(* PLC project VoltPilot-Vorlage PV, VoltPilot VoltPilot EMS 1.0 *)
(* stored: creationDateTime 2026-11-20T00:00:00 *)

(* VoltPilot-Bibliothek · Datentypen des Bausteins Erzeuger-Bild Das Anlagenprogramm füllt diese Strukturen in den Einheiten der Felder des Vertrags docs/contracts/v2/erzeuger-registerbild.md (W, kW, 0,1 %, 0,001, 0,1 kWh, s) und rechnet keine Register: das tut FB_VP_ErzeugerBild. Ein Wert ohne deckendes Gültigkeitsbit hat ein eigenes Feld ...Bekannt: FALSE heißt "kein Wert", der Baustein schreibt dann das Typ-Maximum (Vertrag §1: ungültig ist nie 0). Ein gedeckter Wert braucht keines: ist sein Gültigkeitsbit FALSE, schreibt der Baustein das Typ-Maximum selbst. Ausnahme ist uiPZehntelProzent (Vertrag §3, Wort 24): ohne gültige Vorgabe steht dort der wirksame Ersatzwert. Das Eingangsregister-Abbild: Bild 0..137, Namen ab 140 (höchstens 140 + 32 + 16 * 10 = 332 Wörter). *)
TYPE T_VP_ErzeugerBild : ARRAY[0..331] OF WORD;
END_TYPE

(* Abschnitt A: Anlage und Netzpunkt (Register 12..21). *)
TYPE ST_VP_ErzeugerAnlage : STRUCT
  xNetzpunktGueltig : BOOL;
  xNetzpunktBerechnet : BOOL;
  xNetzpunktTot : BOOL;
  xErzeugungGueltig : BOOL;
  xGasspeicherGueltig : BOOL;
  xGueltigBekannt : BOOL := TRUE;
  uiAlterS : UINT;
  xAlterBekannt : BOOL := TRUE;
  diPNetzpunktW : DINT;
  diPErzeugungW : DINT;
  uiZustand : UINT;
  xZustandBekannt : BOOL := TRUE;
  xNotAus : BOOL;
  xNaSchutz : BOOL;
  xSammelstoerung : BOOL;
  xHandOrt : BOOL;
  xWartung : BOOL;
  xBitsBekannt : BOOL := TRUE;
  uiSpeicherZehntelProzent : UINT;
  uiInstalliertKw : UINT;
  xInstalliertBekannt : BOOL := TRUE;
END_STRUCT;
END_TYPE

(* Abschnitt N: Netzbetreiber (Register 22..27). *)
TYPE ST_VP_ErzeugerNetzbetreiber : STRUCT
  uiKanal : UINT;
  xKanalBekannt : BOOL := TRUE;
  xVorgabeGueltig : BOOL;
  xVerbindungSteht : BOOL;
  xWirkleistungBegrenzt : BOOL;
  xNotAus : BOOL;
  xCosPhiVorgabe : BOOL;
  xKennlinie : BOOL;
  xBitsBekannt : BOOL := TRUE;
  uiPZehntelProzent : UINT;
  xPBekannt : BOOL := TRUE;
  iCosPhiTausendstel : INT;
  uiSeitS : UINT;
  xSeitBekannt : BOOL := TRUE;
  uiZaehler : UINT;
END_STRUCT;
END_TYPE

(* Abschnitt D: Direktvermarkter (Register 28..33). *)
TYPE ST_VP_ErzeugerDirektvermarkter : STRUCT
  uiKanal : UINT;
  xKanalBekannt : BOOL := TRUE;
  xAbschnittGueltig : BOOL;
  xAktivierung : BOOL;
  xStopp : BOOL;
  xBereitGemeldet : BOOL;
  xAktivGemeldet : BOOL;
  xBitsBekannt : BOOL := TRUE;
  udiSollW : UDINT;
  uiSeitS : UINT;
  uiZaehler : UINT;
END_STRUCT;
END_TYPE

(* Abschnitt S: Wirkung (Register 34..37). *)
TYPE ST_VP_ErzeugerWirkung : STRUCT
  xGueltig : BOOL;
  xAnlageFolgt : BOOL;
  xBitsBekannt : BOOL := TRUE;
  uiQuelle : UINT;
  udiGrenzeW : UDINT;
END_STRUCT;
END_TYPE

(* Abschnitt T: eine Einheit (Wechselrichter oder BHKW-Motor), 10 Wörter ab 38 + (n - 1) * 10. *)
TYPE ST_VP_ErzeugerEinheit : STRUCT
  xWerteGueltig : BOOL;
  xSollwertGueltig : BOOL;
  xDvBereit : BOOL;
  xDvAktiv : BOOL;
  xGrundStoerung : BOOL;
  xGrundNetzbetreiber : BOOL;
  xGrundHandOrt : BOOL;
  xGrundWartung : BOOL;
  xGrundGasspeicherLeer : BOOL;
  xGrundSonstiger : BOOL;
  xBitsBekannt : BOOL := TRUE;
  uiZustand : UINT;
  uiArt : UINT;
  xArtBekannt : BOOL := TRUE;
  uiNennKw : UINT;
  xNennBekannt : BOOL := TRUE;
  diPIstW : DINT;
  udiPSollW : UDINT;
  udiEZehntelKwh : UDINT;
  sTyp : STRING(32);
END_STRUCT;
END_TYPE

(* VoltPilot-Bibliothek · Datentypen des Koppelbilds (docs/contracts/v2/koppelbild.md) Das Anlagenprogramm sieht keine Register: es trägt je Stellplatz ein Angebot ein, liest den Wunsch am Ausgang des Bausteins und meldet zurück, was es wirklich anwendet. Codes (Vertrag §7): Art 0 keiner, 1 limit_w (W), 2 limit_pct (0,1 %), 3 setpoint_w (W, Speicher + lädt), 4 on_off (0/1), 5 mode (1..8), 6 setpoint_c (0,1 °C) Ziel 1 erzeugung_gesamt, 2 erzeugungseinheit, 3 speicher, 4 verbraucher, 5 netzbezug, 6 einspeisung, 7 probe Grund 0 keiner, 1 markt, 2 netz, 3 regel, 4 hand, 5 test, 6 vertrag (Nebenversion 1.1; Auskunft, keine Weiche: der Baustein reicht ihn unverändert durch) Abschnitt W: liegt auf den Halteregistern 0..63 des Modbus-TCP-Servers; nur die Edge schreibt. *)
TYPE T_VP_KoppelWunsch : ARRAY[0..63] OF WORD;
END_TYPE

(* Abschnitt Q: liegt auf den Eingangsregistern 1000..1115; nur der Baustein schreibt. *)
TYPE T_VP_KoppelQuittung : ARRAY[0..115] OF WORD;
END_TYPE

(* Was ein Stellplatz anbietet. uiArt 0 = Platz leer. Band in den Einheiten der Art. *)
TYPE ST_VP_Angebot : STRUCT
  uiArt : UINT;
  uiZiel : UINT;
  uiNr : UINT;
  diMin : DINT;
  diMax : DINT;
  xBereit : BOOL;
  xGrundStoerung : BOOL;
  xGrundHandOrt : BOOL;
  xGrundWartung : BOOL;
  xGrundVorrang : BOOL;
  xGrundSonstiger : BOOL;
END_STRUCT;
END_TYPE

(* Was das Anlagenprogramm für das Ziel eines Stellplatzes gerade anwendet, gleich woher es kommt. *)
TYPE ST_VP_Rueckmeldung : STRUCT
  diWirksam : DINT;
  xWirksamBekannt : BOOL;
  xUeberstimmt : BOOL;
END_STRUCT;
END_TYPE

(* Der zugelassene Wunsch eines Stellplatzes. Ohne xGilt fährt das Anlagenprogramm mit eigenen Werten. *)
TYPE ST_VP_Wunsch : STRUCT
  xGilt : BOOL;
  diWert : DINT;
  uiGrund : UINT;
  uiUrteil : UINT;
END_STRUCT;
END_TYPE

(* VoltPilot-Bibliothek · Datentypen des Bausteins WAGO-Bild (Energiekarten) Das Anlagenprogramm kopiert je 3-Phasen-Leistungsmessklemme 750-494/-495 („Energiekarte“) die Werte, die es aus der Karte gelesen hat, in eine ST_VP_WagoKarte - unverändert, in der Skalierung der Karte (docs/contracts/v2/wago-registerbild.md §4). Umgerechnet wird nichts: Einheit, Faktor und Vorzeichen kommen aus dem Katalog und dem Hardwareblatt der Anlage. Jeder Teil hat sein Feld ...Gelesen: FALSE heißt "dieser Teil ist unbekannt", der Baustein löscht dann das Gültigkeitsbit und schreibt das Typ-Maximum - nie 0, nie einen alten Wert. Das Abbild: Kopf 12 Wörter und höchstens 16 Karten zu je 42 Wörtern (12 + 16 * 42 = 684). *)
TYPE T_VP_WagoBild : ARRAY[0..683] OF WORD;
END_TYPE

(* Eine Energiekarte (Vertrag §4). *)
TYPE ST_VP_WagoKarte : STRUCT
  uiSteckplatz : UINT;
  uiKartentyp : UINT;
  uiVariante : UINT;
  xKarteGelesen : BOOL;
  xKr32Gelesen : BOOL;
  wKr32 : WORD;
  xKr35Gelesen : BOOL;
  wKr35 : WORD;
  xStatusGelesen : BOOL;
  awStatus : ARRAY[0..11] OF WORD;
  adwMesswert : ARRAY[1..12] OF DWORD;
END_STRUCT;
END_TYPE

VAR_GLOBAL  (* GVL_VoltPilot *)
  aErzeugerBild : T_VP_ErzeugerBild;
  aKoppelQuittung : T_VP_KoppelQuittung;
  aKoppelWunsch : T_VP_KoppelWunsch;
  aWagoBild : T_VP_WagoBild;
  xProbeLampe : BOOL;
END_VAR

(* VoltPilot-Bibliothek · Baustein Erzeuger-Bild Füllt das "VoltPilot-Registerbild Erzeuger v1" (schlanke Fassung 1.0, docs/contracts/v2/erzeuger-registerbild.md) aus den getippten Werten des Anlagenprogramms. Das Abbild aBild liegt auf den Eingangsregistern des Modbus-TCP-Servers ab Adresse 0 (Funktionscode 4); die Box liest es alle 5 s, auf einem PFC200 mit VoltPilot über 127.0.0.1. Aufruf: einmal je Zyklus in der Task, die das Abbild auch dem Modbus-Server übergibt. fbBild(uiProgrammstand := 2611, uiAnlagenart := 1, uiTeAnzahl := 3, stAnlage := stAnlage, stNetzbetreiber := stNb, stDirektvermarkter := stDv, stWirkung := stWirkung, astEinheit := astEinheit, xMitNamen := TRUE, sNetzbetreiber := 'Netzbetreiber', sDirektvermarkter := '', aBild := GVL_VoltPilot.aErzeugerBild); Was der Baustein selbst hält: - Kopf: Signatur, Prüfwert, Fassung 1.0 - feste Werte, der Prüfwert über VP_SetzeU32; - Herzschlag: +1 je Sekunde seit Programmstart, 65535 -> 0 (Vertrag §8); bleibt der Aufruf aus, steht er, und die Box hält alle Werte nach drei gleichen Lesungen für veraltet; - Typ-Maximum für jeden gedeckten Wert, dessen Gültigkeitsbit fehlt; - Wörter von Einheiten über uiTeAnzahl hinaus und ohne Namen den Namenbereich auf 0. Grenzen: höchstens 10 Einheiten; uiTeAnzahl 0 oder über 10 schreibt der Baustein, wie er sie bekommt - die Box liest das Bild dann nicht (te_anzahl_ungueltig), sieht aber Kopf und Herzschlag (so meldet sich das Grundprogramm ohne Anlage). *)
FUNCTION_BLOCK FB_VP_ErzeugerBild
  VAR_INPUT
    udiSteuerungId : UDINT := 16#FFFFFFFF;
    uiProgrammstand : UINT := 16#FFFF;
    uiAnlagenart : UINT := 16#FFFF;
    uiTeAnzahl : UINT;
    stAnlage : ST_VP_ErzeugerAnlage;
    stNetzbetreiber : ST_VP_ErzeugerNetzbetreiber;
    stDirektvermarkter : ST_VP_ErzeugerDirektvermarkter;
    stWirkung : ST_VP_ErzeugerWirkung;
    astEinheit : ARRAY[1..10] OF ST_VP_ErzeugerEinheit;
    xMitNamen : BOOL;
    sNetzbetreiber : STRING(32);
    sDirektvermarkter : STRING(32);
  END_VAR
  VAR_IN_OUT
    aBild : T_VP_ErzeugerBild;
  END_VAR
  VAR
    uiHerzschlag : UINT;
    xGestartet : BOOL;
    tLetzte : TIME;
    tJetzt : TIME;
    udiSekunden : UDINT;
    n : UINT;
    uiBasis : UINT;
    i : UINT;
    wBits : WORD;
  END_VAR

(* --- Herzschlag: +1 je Sekunde, beim Programmstart 0, 65535 -> 0 ---------------------------- *)
tJetzt := TIME();
IF NOT xGestartet THEN
    tLetzte := tJetzt;
    xGestartet := TRUE;
END_IF
udiSekunden := TIME_TO_UDINT(tJetzt - tLetzte) / 1000;
IF udiSekunden > 0 THEN
    uiHerzschlag := uiHerzschlag + UDINT_TO_UINT(udiSekunden AND 16#FFFF);
    tLetzte := tLetzte + UDINT_TO_TIME(udiSekunden * 1000);
END_IF

(* --- Kopf (0..11) ------------------------------------------------------------------------- *)
aBild[0] := 16#5650;   (* "VP" *)
aBild[1] := 16#455A;   (* "EZ" *)
VP_SetzeU32(aBild := aBild, uiAdresse := 2, udiWert := 16#01020304, xBekannt := TRUE);
aBild[4] := 16#0100;   (* Fassung 1.0 *)
aBild[5] := UINT_TO_WORD(uiTeAnzahl);
aBild[6] := UINT_TO_WORD(uiHerzschlag);
aBild[7] := UINT_TO_WORD(uiProgrammstand);
VP_SetzeU32(aBild := aBild, uiAdresse := 8, udiWert := udiSteuerungId, xBekannt := TRUE);
aBild[10] := UINT_TO_WORD(uiAnlagenart);
IF xMitNamen THEN
    aBild[11] := 140;
ELSE
    aBild[11] := 0;
END_IF

(* --- A: Anlage und Netzpunkt (12..21) ------------------------------------------------------ *)
wBits := VP_Bit(stAnlage.xNetzpunktGueltig, 0) OR VP_Bit(stAnlage.xNetzpunktBerechnet, 1)
    OR VP_Bit(stAnlage.xNetzpunktTot, 2) OR VP_Bit(stAnlage.xErzeugungGueltig, 3)
    OR VP_Bit(stAnlage.xGasspeicherGueltig, 4);
VP_SetzeU16(aBild := aBild, uiAdresse := 12, uiWert := WORD_TO_UINT(wBits), xBekannt := stAnlage.xGueltigBekannt);
VP_SetzeU16(aBild := aBild, uiAdresse := 13, uiWert := stAnlage.uiAlterS, xBekannt := stAnlage.xAlterBekannt);
VP_SetzeS32(aBild := aBild, uiAdresse := 14, diWert := stAnlage.diPNetzpunktW,
    xBekannt := stAnlage.xGueltigBekannt AND stAnlage.xNetzpunktGueltig);
VP_SetzeS32(aBild := aBild, uiAdresse := 16, diWert := stAnlage.diPErzeugungW,
    xBekannt := stAnlage.xGueltigBekannt AND stAnlage.xErzeugungGueltig);
VP_SetzeU16(aBild := aBild, uiAdresse := 18, uiWert := stAnlage.uiZustand, xBekannt := stAnlage.xZustandBekannt);
wBits := VP_Bit(stAnlage.xNotAus, 0) OR VP_Bit(stAnlage.xNaSchutz, 1) OR VP_Bit(stAnlage.xSammelstoerung, 2)
    OR VP_Bit(stAnlage.xHandOrt, 3) OR VP_Bit(stAnlage.xWartung, 4);
VP_SetzeU16(aBild := aBild, uiAdresse := 19, uiWert := WORD_TO_UINT(wBits), xBekannt := stAnlage.xBitsBekannt);
VP_SetzeU16(aBild := aBild, uiAdresse := 20, uiWert := stAnlage.uiSpeicherZehntelProzent,
    xBekannt := stAnlage.xGueltigBekannt AND stAnlage.xGasspeicherGueltig);
VP_SetzeU16(aBild := aBild, uiAdresse := 21, uiWert := stAnlage.uiInstalliertKw, xBekannt := stAnlage.xInstalliertBekannt);

(* --- N: Netzbetreiber (22..27) ------------------------------------------------------------- *)
VP_SetzeU16(aBild := aBild, uiAdresse := 22, uiWert := stNetzbetreiber.uiKanal, xBekannt := stNetzbetreiber.xKanalBekannt);
wBits := VP_Bit(stNetzbetreiber.xVorgabeGueltig, 0) OR VP_Bit(stNetzbetreiber.xVerbindungSteht, 1)
    OR VP_Bit(stNetzbetreiber.xWirkleistungBegrenzt, 2) OR VP_Bit(stNetzbetreiber.xNotAus, 3)
    OR VP_Bit(stNetzbetreiber.xCosPhiVorgabe, 4) OR VP_Bit(stNetzbetreiber.xKennlinie, 5);
VP_SetzeU16(aBild := aBild, uiAdresse := 23, uiWert := WORD_TO_UINT(wBits), xBekannt := stNetzbetreiber.xBitsBekannt);
(* Wort 24 ohne gültige Vorgabe: der wirksame Ersatzwert, nicht das Typ-Maximum (Vertrag §3) *)
VP_SetzeU16(aBild := aBild, uiAdresse := 24, uiWert := stNetzbetreiber.uiPZehntelProzent, xBekannt := stNetzbetreiber.xPBekannt);
VP_SetzeS16(aBild := aBild, uiAdresse := 25, iWert := stNetzbetreiber.iCosPhiTausendstel,
    xBekannt := stNetzbetreiber.xBitsBekannt AND stNetzbetreiber.xVorgabeGueltig);
VP_SetzeU16(aBild := aBild, uiAdresse := 26, uiWert := stNetzbetreiber.uiSeitS, xBekannt := stNetzbetreiber.xSeitBekannt);
aBild[27] := UINT_TO_WORD(stNetzbetreiber.uiZaehler);

(* --- D: Direktvermarkter (28..33) ---------------------------------------------------------- *)
VP_SetzeU16(aBild := aBild, uiAdresse := 28, uiWert := stDirektvermarkter.uiKanal, xBekannt := stDirektvermarkter.xKanalBekannt);
wBits := VP_Bit(stDirektvermarkter.xAbschnittGueltig, 0) OR VP_Bit(stDirektvermarkter.xAktivierung, 1)
    OR VP_Bit(stDirektvermarkter.xStopp, 2) OR VP_Bit(stDirektvermarkter.xBereitGemeldet, 3)
    OR VP_Bit(stDirektvermarkter.xAktivGemeldet, 4);
VP_SetzeU16(aBild := aBild, uiAdresse := 29, uiWert := WORD_TO_UINT(wBits), xBekannt := stDirektvermarkter.xBitsBekannt);
VP_SetzeU32(aBild := aBild, uiAdresse := 30, udiWert := stDirektvermarkter.udiSollW,
    xBekannt := stDirektvermarkter.xBitsBekannt AND stDirektvermarkter.xAbschnittGueltig);
VP_SetzeU16(aBild := aBild, uiAdresse := 32, uiWert := stDirektvermarkter.uiSeitS,
    xBekannt := stDirektvermarkter.xBitsBekannt AND stDirektvermarkter.xAbschnittGueltig);
(* d_zaehler hat keinen Ungültig-Wert; ohne gültigen Abschnitt liest ihn die Box nicht *)
aBild[33] := UINT_TO_WORD(stDirektvermarkter.uiZaehler);

(* --- S: Wirkung (34..37) ------------------------------------------------------------------- *)
VP_SetzeU16(aBild := aBild, uiAdresse := 34, uiWert := stWirkung.uiQuelle,
    xBekannt := stWirkung.xBitsBekannt AND stWirkung.xGueltig);
wBits := VP_Bit(stWirkung.xGueltig, 0) OR VP_Bit(stWirkung.xAnlageFolgt, 1);
VP_SetzeU16(aBild := aBild, uiAdresse := 35, uiWert := WORD_TO_UINT(wBits), xBekannt := stWirkung.xBitsBekannt);
VP_SetzeU32(aBild := aBild, uiAdresse := 36, udiWert := stWirkung.udiGrenzeW,
    xBekannt := stWirkung.xBitsBekannt AND stWirkung.xGueltig);

(* --- T: je Einheit 10 Wörter ab 38 + (n - 1) * 10 ------------------------------------------ *)
FOR n := 1 TO 10 DO
    uiBasis := 38 + (n - 1) * 10;
    IF n <= uiTeAnzahl THEN
        VP_SetzeU16(aBild := aBild, uiAdresse := uiBasis, uiWert := astEinheit[n].uiZustand,
            xBekannt := astEinheit[n].xBitsBekannt AND astEinheit[n].xWerteGueltig);
        wBits := VP_Bit(astEinheit[n].xWerteGueltig, 0) OR VP_Bit(astEinheit[n].xSollwertGueltig, 1)
            OR VP_Bit(astEinheit[n].xDvBereit, 2) OR VP_Bit(astEinheit[n].xDvAktiv, 3)
            OR VP_Bit(astEinheit[n].xGrundStoerung, 4) OR VP_Bit(astEinheit[n].xGrundNetzbetreiber, 5)
            OR VP_Bit(astEinheit[n].xGrundHandOrt, 6) OR VP_Bit(astEinheit[n].xGrundWartung, 7)
            OR VP_Bit(astEinheit[n].xGrundGasspeicherLeer, 8) OR VP_Bit(astEinheit[n].xGrundSonstiger, 9);
        VP_SetzeU16(aBild := aBild, uiAdresse := uiBasis + 1, uiWert := WORD_TO_UINT(wBits),
            xBekannt := astEinheit[n].xBitsBekannt);
        VP_SetzeU16(aBild := aBild, uiAdresse := uiBasis + 2, uiWert := astEinheit[n].uiArt,
            xBekannt := astEinheit[n].xArtBekannt);
        VP_SetzeU16(aBild := aBild, uiAdresse := uiBasis + 3, uiWert := astEinheit[n].uiNennKw,
            xBekannt := astEinheit[n].xNennBekannt);
        VP_SetzeS32(aBild := aBild, uiAdresse := uiBasis + 4, diWert := astEinheit[n].diPIstW,
            xBekannt := astEinheit[n].xBitsBekannt AND astEinheit[n].xWerteGueltig);
        VP_SetzeU32(aBild := aBild, uiAdresse := uiBasis + 6, udiWert := astEinheit[n].udiPSollW,
            xBekannt := astEinheit[n].xBitsBekannt AND astEinheit[n].xSollwertGueltig);
        VP_SetzeU32(aBild := aBild, uiAdresse := uiBasis + 8, udiWert := astEinheit[n].udiEZehntelKwh,
            xBekannt := astEinheit[n].xBitsBekannt AND astEinheit[n].xWerteGueltig);
    ELSE
        (* frei: nichts Altes aus einer früheren Zahl der Einheiten bleibt stehen *)
        FOR i := uiBasis TO uiBasis + 9 DO
            aBild[i] := 0;
        END_FOR
    END_IF
END_FOR
FOR i := 138 TO 139 DO
    aBild[i] := 0;
END_FOR

(* --- Namen ab 140: Netzbetreiber +0, Direktvermarkter +16, Typ der Einheit n +32 + (n - 1) * 16 *)
IF xMitNamen THEN
    VP_SetzeText(aBild := aBild, uiAdresse := 140, sText := sNetzbetreiber);
    VP_SetzeText(aBild := aBild, uiAdresse := 156, sText := sDirektvermarkter);
    FOR n := 1 TO 10 DO
        IF n <= uiTeAnzahl THEN
            VP_SetzeText(aBild := aBild, uiAdresse := 172 + (n - 1) * 16, sText := astEinheit[n].sTyp);
        ELSE
            VP_SetzeText(aBild := aBild, uiAdresse := 172 + (n - 1) * 16, sText := '');
        END_IF
    END_FOR
ELSE
    FOR i := 140 TO 331 DO
        aBild[i] := 0;
    END_FOR
END_IF
END_FUNCTION_BLOCK

(* VoltPilot-Bibliothek · Baustein Koppelbild Die SPS-Seite des "VoltPilot-Koppelbild v1" (docs/contracts/v2/koppelbild.md): die Edge schreibt Wünsche in die Halteregister 0..63, der Baustein prüft sie, begrenzt jeden auf das Angebot und reicht ihn dem Anlagenprogramm; die Quittung steht in den Eingangsregistern 1000..1115. Die SPS entscheidet immer selbst: ein Wunsch ist nie ein Befehl. Aufruf: einmal je Zyklus in der Task, die die Abbilder auch dem Modbus-Server übergibt. fbKoppel(udiSteuerungId := 1042, xFernsteuerungFrei := xSchluesselFern, xHandOrt := xHand, aAngebot := aAngebot, aRueckmeldung := aRueck, aWunschRegister := GVL_VoltPilot.aKoppelWunsch, aQuittungRegister := GVL_VoltPilot.aKoppelQuittung); IF fbKoppel.aWunsch[1].xGilt THEN diGrenze := MIN(diGrenze, fbKoppel.aWunsch[1].diWert); END_IF Was der Baustein selbst hält: - jeder Wunsch läuft von selbst ab: höchstens frist_s ab Empfang, nie länger als tHoechsteFrist (Vorgabe 60 s); fällt die Edge aus, fährt die Anlage danach mit eigenen Werten; - Lebenszeichen: Herzschlag +1 je Sekunde (wie im Erzeuger-Bild), edge_lebt aus dem letzten gültigen Telegramm; - geprüft wird nur ein Telegramm, dessen Wörter sich geändert haben, in der Reihenfolge von Vertrag §5; ein abgelehntes bewirkt nichts, das vorige gilt bis zu seiner Frist; - Hand/Ort nimmt jedem Stellplatz die Bereitschaft; ohne Fernsteuerung gilt kein Wunsch. Was beim ersten Aufruf in den Halteregistern steht, ist kein Telegramm, nur der Vergleichsstand. *)
FUNCTION_BLOCK FB_VP_Koppelbild
  VAR_INPUT
    udiSteuerungId : UDINT;
    xFernsteuerungFrei : BOOL;
    xHandOrt : BOOL;
    aAngebot : ARRAY[1..8] OF ST_VP_Angebot;
    aRueckmeldung : ARRAY[1..8] OF ST_VP_Rueckmeldung;
    tHoechsteFrist : TIME := T#60S;
    uiBibliothek : UINT := 16#0100;
  END_VAR
  VAR_OUTPUT
    aWunsch : ARRAY[1..8] OF ST_VP_Wunsch;
    xEdgeLebt : BOOL;
    uiKopfUrteil : UINT;
    uiRestS : UINT;
  END_VAR
  VAR_IN_OUT
    aWunschRegister : T_VP_KoppelWunsch;
    aQuittungRegister : T_VP_KoppelQuittung;
  END_VAR
  VAR
    uiHerzschlag : UINT;
    xGestartet : BOOL;
    tLetzte : TIME;
    tJetzt : TIME;
    udiSekunden : UDINT;
    xErster : BOOL := TRUE;
    aLetzte : T_VP_KoppelWunsch;
    aGilt : T_VP_KoppelWunsch;
    xHatTelegramm : BOOL;
    xFristLaeuft : BOOL;
    uiOhneFrist : UINT;
    tAnnahme : TIME;
    udiFristMs : UDINT;
    udiSeitMs : UDINT;
    xLebt : BOOL;
    uiQSitzung : UINT;
    uiQHerzschlag : UINT;
    uiAngenommen : UINT;
    uiAbgelehnt : UINT;
    xGeaendert : BOOL;
    uiGrund : UINT;
    udiFrist : UDINT;
    i : UINT;
    n : UINT;
    uiW : UINT;
    uiQ : UINT;
    uiAnzahl : UINT;
    xLeer : BOOL;
    xBereit : BOOL;
    uiArtW : UINT;
    diW : DINT;
    diWert : DINT;
    uiUrteil : UINT;
  END_VAR

(* --- Herzschlag: +1 je Sekunde seit Programmstart, 65535 -> 0 ------------------------------ *)
tJetzt := TIME();
IF NOT xGestartet THEN
    tLetzte := tJetzt;
    xGestartet := TRUE;
END_IF
udiSekunden := TIME_TO_UDINT(tJetzt - tLetzte) / 1000;
IF udiSekunden > 0 THEN
    uiHerzschlag := uiHerzschlag + UDINT_TO_UINT(udiSekunden AND 16#FFFF);
    tLetzte := tLetzte + UDINT_TO_TIME(udiSekunden * 1000);
END_IF

(* --- Telegramm prüfen, wenn sich ein Wort geändert hat (Vertrag §5) ------------------------- *)
IF xErster THEN
    aLetzte := aWunschRegister;
    xErster := FALSE;
ELSE
    xGeaendert := FALSE;
    FOR i := 0 TO 63 DO
        IF aWunschRegister[i] <> aLetzte[i] THEN
            xGeaendert := TRUE;
        END_IF
    END_FOR
    IF xGeaendert THEN
        aLetzte := aWunschRegister;
        udiFrist := WORD_TO_UDINT(aWunschRegister[10]);
        uiGrund := 0;
        IF aWunschRegister[0] <> 16#5650 OR aWunschRegister[1] <> 16#4B57 THEN
            uiGrund := 2;
        ELSIF SHR(aWunschRegister[4], 8) <> 1 THEN
            uiGrund := 3;
        ELSIF aWunschRegister[2] <> 16#0102 OR aWunschRegister[3] <> 16#0304 THEN
            uiGrund := 4;
        ELSIF VP_KoppelSiegelW(aW := aWunschRegister) <> aWunschRegister[15] THEN
            uiGrund := 5;
        ELSIF VP_KoppelLiesU32(aW := aWunschRegister, uiAdresse := 8) <> udiSteuerungId THEN
            uiGrund := 6;
        ELSIF udiFrist < 5 OR udiFrist > 600 OR aWunschRegister[6] = 0 OR aWunschRegister[6] = 16#FFFF
                OR aWunschRegister[5] <> 8 THEN
            uiGrund := 7;
        END_IF
        IF uiGrund <> 0 THEN
            (* dieses Telegramm bewirkt nichts; das vorige gilt bis zu seiner Frist *)
            uiAbgelehnt := uiAbgelehnt + 1;
            uiKopfUrteil := uiGrund;
        ELSE
            aGilt := aWunschRegister;
            xHatTelegramm := TRUE;
            uiQSitzung := WORD_TO_UINT(aWunschRegister[6]);
            uiQHerzschlag := WORD_TO_UINT(aWunschRegister[7]);
            uiAngenommen := uiAngenommen + 1;
            tAnnahme := tJetzt;
            xLebt := TRUE;
            IF xFernsteuerungFrei THEN
                udiFristMs := MIN(udiFrist * 1000, TIME_TO_UDINT(tHoechsteFrist));
                xFristLaeuft := TRUE;
                uiKopfUrteil := 1;
            ELSE
                xFristLaeuft := FALSE;
                uiOhneFrist := 2;
                uiKopfUrteil := 9;
            END_IF
        END_IF
    END_IF
END_IF

(* --- Fernsteuerung entzogen: alle Wünsche fallen sofort ------------------------------------ *)
IF NOT xFernsteuerungFrei AND xFristLaeuft THEN
    xFristLaeuft := FALSE;
    uiOhneFrist := 2;
    uiKopfUrteil := 9;
END_IF

(* --- Frist: läuft von selbst ab ------------------------------------------------------------ *)
udiSeitMs := TIME_TO_UDINT(tJetzt - tAnnahme);
IF xFristLaeuft AND udiSeitMs >= udiFristMs THEN
    xFristLaeuft := FALSE;
    uiOhneFrist := 1;
    uiKopfUrteil := 8;
END_IF
IF xFristLaeuft THEN
    uiRestS := UDINT_TO_UINT((udiFristMs - udiSeitMs + 999) / 1000);
ELSE
    uiRestS := 0;
END_IF
(* einmal still, bleibt still: auch wenn TIME() nach 49 Tagen überläuft *)
IF xLebt AND udiSeitMs >= 15000 THEN
    xLebt := FALSE;
END_IF
xEdgeLebt := xLebt;

(* --- Kopf der Quittung (1000..1019, hier 0..19) -------------------------------------------- *)
aQuittungRegister[0] := 16#5650;   (* "VP" *)
aQuittungRegister[1] := 16#4B51;   (* "KQ" *)
VP_KoppelSetzeU32(aQ := aQuittungRegister, uiAdresse := 2, udiWert := 16#01020304);
aQuittungRegister[4] := 16#0100;   (* Fassung 1.0 *)
aQuittungRegister[6] := UINT_TO_WORD(uiHerzschlag);
aQuittungRegister[7] := UINT_TO_WORD(uiBibliothek);
VP_KoppelSetzeU32(aQ := aQuittungRegister, uiAdresse := 8, udiWert := udiSteuerungId);
aQuittungRegister[10] := UINT_TO_WORD(uiKopfUrteil);
aQuittungRegister[11] := UINT_TO_WORD(uiQSitzung);
aQuittungRegister[12] := UINT_TO_WORD(uiQHerzschlag);
aQuittungRegister[13] := UINT_TO_WORD(uiRestS);
aQuittungRegister[14] := VP_Bit(xGesetzt := xFernsteuerungFrei, uiBit := 0)
    OR VP_Bit(xGesetzt := xLebt, uiBit := 1) OR VP_Bit(xGesetzt := xHandOrt, uiBit := 2);
aQuittungRegister[15] := UINT_TO_WORD(uiAngenommen);
aQuittungRegister[16] := UINT_TO_WORD(uiAbgelehnt);
aQuittungRegister[17] := 0;
aQuittungRegister[18] := 0;

(* --- je Stellplatz: Angebot, Urteil, zugelassener Wert, wirksam (Vertrag §5) ---------------- *)
uiAnzahl := 0;
FOR n := 1 TO 8 DO
    uiW := 16 + (n - 1) * 6;
    uiQ := 20 + (n - 1) * 12;
    xLeer := aAngebot[n].uiArt = 0;
    xBereit := NOT xLeer AND aAngebot[n].xBereit AND NOT xHandOrt;
    uiUrteil := 0;
    diWert := 0;
    aWunsch[n].xGilt := FALSE;
    aWunsch[n].uiGrund := 0;
    IF NOT xLeer THEN
        uiAnzahl := uiAnzahl + 1;
    END_IF
    IF xHatTelegramm THEN
        uiArtW := WORD_TO_UINT(aGilt[uiW]);
        diW := UDINT_TO_DINT(SHL(WORD_TO_UDINT(aGilt[uiW + 2]), 16) OR WORD_TO_UDINT(aGilt[uiW + 3]));
        IF NOT xFristLaeuft THEN
            IF uiArtW <> 0 AND uiOhneFrist = 1 THEN
                uiUrteil := 7;
            ELSIF uiArtW <> 0 AND uiOhneFrist = 2 THEN
                uiUrteil := 5;
            END_IF
        ELSIF uiArtW = 0 THEN
            uiUrteil := 0;
        ELSIF xLeer OR uiArtW <> aAngebot[n].uiArt THEN
            uiUrteil := 3;
        ELSIF diW = 16#7FFFFFFF THEN
            uiUrteil := 4;
        ELSIF NOT xBereit THEN
            uiUrteil := 5;
        ELSE
            diWert := LIMIT(aAngebot[n].diMin, diW, aAngebot[n].diMax);
            IF aRueckmeldung[n].xUeberstimmt THEN
                uiUrteil := 6;
            ELSIF diWert <> diW THEN
                uiUrteil := 2;
            ELSE
                uiUrteil := 1;
            END_IF
            aWunsch[n].xGilt := TRUE;
            aWunsch[n].uiGrund := WORD_TO_UINT(aGilt[uiW + 1]);
        END_IF
        aQuittungRegister[uiQ + 9] := aGilt[uiW + 4];
    ELSE
        aQuittungRegister[uiQ + 9] := 0;
    END_IF
    aWunsch[n].diWert := diWert;
    aWunsch[n].uiUrteil := uiUrteil;
    aQuittungRegister[uiQ] := UINT_TO_WORD(aAngebot[n].uiArt);
    IF xLeer THEN
        aQuittungRegister[uiQ + 1] := 0;
        aQuittungRegister[uiQ + 2] := 0;
        aQuittungRegister[uiQ + 3] := 0;
    ELSE
        aQuittungRegister[uiQ + 1] := UINT_TO_WORD(aAngebot[n].uiZiel);
        aQuittungRegister[uiQ + 2] := UINT_TO_WORD(aAngebot[n].uiNr);
        aQuittungRegister[uiQ + 3] := VP_Bit(xGesetzt := xBereit, uiBit := 0)
            OR VP_Bit(xGesetzt := aAngebot[n].xGrundStoerung, uiBit := 1)
            OR VP_Bit(xGesetzt := aAngebot[n].xGrundHandOrt OR xHandOrt, uiBit := 2)
            OR VP_Bit(xGesetzt := aAngebot[n].xGrundWartung, uiBit := 3)
            OR VP_Bit(xGesetzt := aAngebot[n].xGrundVorrang, uiBit := 4)
            OR VP_Bit(xGesetzt := aAngebot[n].xGrundSonstiger, uiBit := 5);
    END_IF
    VP_KoppelSetzeS32(aQ := aQuittungRegister, uiAdresse := uiQ + 4, diWert := aAngebot[n].diMin, xBekannt := NOT xLeer);
    VP_KoppelSetzeS32(aQ := aQuittungRegister, uiAdresse := uiQ + 6, diWert := aAngebot[n].diMax, xBekannt := NOT xLeer);
    aQuittungRegister[uiQ + 8] := UINT_TO_WORD(uiUrteil);
    VP_KoppelSetzeS32(aQ := aQuittungRegister, uiAdresse := uiQ + 10, diWert := aRueckmeldung[n].diWirksam,
        xBekannt := aRueckmeldung[n].xWirksamBekannt);
END_FOR
aQuittungRegister[5] := UINT_TO_WORD(uiAnzahl);
aQuittungRegister[19] := VP_KoppelSiegelQ(aQ := aQuittungRegister);
END_FUNCTION_BLOCK

(* VoltPilot-Bibliothek · Baustein WAGO-Bild (Energiekarten) Füllt das "VoltPilot-Registerbild WAGO v1" (Fassung 1.0, docs/contracts/v2/wago-registerbild.md) aus den Werten der 3-Phasen-Leistungsmessklemmen 750-494/-495, die das Anlagenprogramm aus den Karten liest: von außen kommt niemand an die Klemmen, ein Programm muss sie kopieren. Das Abbild aBild liegt auf den Registern des Modbus-TCP-Servers ab der Basisadresse der Anlage; für eine neue Anlage auf einem PFC200 mit VoltPilot sind das die Eingangsregister ab 2000 (Funktionscode 4), neben dem Erzeuger-Bild ab 0. Aufruf: einmal je Zyklus in der Task, die das Abbild auch dem Modbus-Server übergibt. fbWago(udiControllerKennung := 1, uiKartenzahl := 2, astKarte := astKarte, aBild := GVL_VoltPilot.aWagoBild); Was der Baustein selbst hält: - Kopf: Signatur "VP" "RB", Fassung 1.0, Längen 12 und 42, der Prüfwert über VP_WagoSetze32; - Herzschlag: +1 je Sekunde seit Programmstart, 65535 -> 0 (Vertrag §3); bleibt der Aufruf aus, steht er, und die Box hält die Kartenwerte nach drei gleichen Lesungen für veraltet; - Gültigkeit: je Karte die Bits aus den Feldern ...Gelesen; ein unbekannter Teil steht als Typ-Maximum im Bild (Int32 16#7FFFFFFF, sonst 16#FFFF bzw. 16#FFFFFFFF), nie als 0; - Wörter von Karten über uiKartenzahl hinaus auf 0. Grenzen: höchstens 16 Karten. uiKartenzahl über 16 schreibt der Baustein, wie er sie bekommt, füllt aber nur 16 Blöcke - die Box liest das Bild dann nicht (Kartenzahl weicht vom Soll ab oder die Register fehlen), statt Karten zu erfinden. *)
FUNCTION_BLOCK FB_VP_WagoBild
  VAR_INPUT
    udiControllerKennung : UDINT;
    xWortfolgeLittle : BOOL;
    uiKartenzahl : UINT;
    astKarte : ARRAY[1..16] OF ST_VP_WagoKarte;
  END_VAR
  VAR_IN_OUT
    aBild : T_VP_WagoBild;
  END_VAR
  VAR
    uiHerzschlag : UINT;
    xGestartet : BOOL;
    tLetzte : TIME;
    tJetzt : TIME;
    udiSekunden : UDINT;
    n : UINT;
    uiBasis : UINT;
    i : UINT;
    wBits : WORD;
    dwUngueltig : DWORD;
  END_VAR

(* --- Herzschlag: +1 je Sekunde, beim Programmstart 0, 65535 -> 0 ---------------------------- *)
tJetzt := TIME();
IF NOT xGestartet THEN
    tLetzte := tJetzt;
    xGestartet := TRUE;
END_IF
udiSekunden := TIME_TO_UDINT(tJetzt - tLetzte) / 1000;
IF udiSekunden > 0 THEN
    uiHerzschlag := uiHerzschlag + UDINT_TO_UINT(udiSekunden AND 16#FFFF);
    tLetzte := tLetzte + UDINT_TO_TIME(udiSekunden * 1000);
END_IF

(* --- Kopf (0..11) ------------------------------------------------------------------------- *)
aBild[0] := 16#5650;   (* "VP" *)
aBild[1] := 16#5242;   (* "RB" *)
aBild[2] := 1;         (* Hauptversion *)
aBild[3] := 0;         (* Nebenversion *)
aBild[4] := 12;        (* Kopflänge *)
aBild[5] := 42;        (* Kartenblocklänge *)
aBild[6] := UINT_TO_WORD(uiKartenzahl);
aBild[7] := UINT_TO_WORD(uiHerzschlag);
VP_WagoSetze32(aBild := aBild, uiAdresse := 8, dwWert := 16#01020304, xLittle := xWortfolgeLittle);
VP_WagoSetze32(aBild := aBild, uiAdresse := 10, dwWert := UDINT_TO_DWORD(udiControllerKennung),
    xLittle := xWortfolgeLittle);

(* --- Karten: Block n beginnt bei 12 + (n - 1) * 42 ------------------------------------------ *)
FOR n := 1 TO 16 DO
    uiBasis := 12 + (n - 1) * 42;
    IF n > uiKartenzahl THEN
        FOR i := 0 TO 41 DO
            aBild[uiBasis + i] := 0;
        END_FOR
    ELSE
        aBild[uiBasis] := UINT_TO_WORD(astKarte[n].uiSteckplatz);
        aBild[uiBasis + 1] := UINT_TO_WORD(astKarte[n].uiKartentyp);
        aBild[uiBasis + 2] := UINT_TO_WORD(astKarte[n].uiVariante);
        wBits := 0;
        IF astKarte[n].xKarteGelesen THEN
            wBits := wBits OR 16#0001;
        END_IF
        IF astKarte[n].xKr32Gelesen THEN
            wBits := wBits OR 16#0002;
        END_IF
        IF astKarte[n].xKr35Gelesen THEN
            wBits := wBits OR 16#0004;
        END_IF
        IF astKarte[n].xStatusGelesen THEN
            wBits := wBits OR 16#0008;
        END_IF
        aBild[uiBasis + 3] := wBits;
        IF astKarte[n].xKr32Gelesen THEN
            aBild[uiBasis + 4] := astKarte[n].wKr32;
        ELSE
            aBild[uiBasis + 4] := 16#FFFF;
        END_IF
        IF astKarte[n].xKr35Gelesen THEN
            aBild[uiBasis + 5] := astKarte[n].wKr35;
        ELSE
            aBild[uiBasis + 5] := 16#FFFF;
        END_IF
        FOR i := 0 TO 11 DO
            IF astKarte[n].xStatusGelesen THEN
                aBild[uiBasis + 6 + i] := astKarte[n].awStatus[i];
            ELSE
                aBild[uiBasis + 6 + i] := 16#FFFF;
            END_IF
        END_FOR
        (* Messwerte ab Offset 18, je zwei Wörter, in der Wortfolge der Anlage *)
        FOR i := 1 TO 12 DO
            IF astKarte[n].xKarteGelesen THEN
                VP_WagoSetze32(aBild := aBild, uiAdresse := uiBasis + 16 + 2 * i,
                    dwWert := astKarte[n].adwMesswert[i], xLittle := xWortfolgeLittle);
            ELSE
                (* ungültig ist das Typ-Maximum des Felds: Wirkleistung L1..L3 sind Int32 *)
                IF i >= 3 AND i <= 5 THEN
                    dwUngueltig := 16#7FFFFFFF;
                ELSE
                    dwUngueltig := 16#FFFFFFFF;
                END_IF
                VP_WagoSetze32(aBild := aBild, uiAdresse := uiBasis + 16 + 2 * i,
                    dwWert := dwUngueltig, xLittle := xWortfolgeLittle);
            END_IF
        END_FOR
    END_IF
END_FOR
END_FUNCTION_BLOCK

(* VoltPilot-Bibliothek · Packfunktionen des Erzeuger-Bilds Jede Zahl geht über genau eine dieser Funktionen ins Bild - auch der Prüfwert 16#01020304 (Vertrag §1, Lesart 9): schriebe das Programm ihn als zwei Konstanten, prüfte er seine Packfunktion nicht, und ein falsch packendes Programm sähe gesund aus (Fall E5). Wortfolge: höherwertiges Wort zuerst. Ungültig: das Typ-Maximum, nie 0. *)
FUNCTION VP_SetzeU16 : BOOL
  VAR_INPUT
    uiAdresse : UINT;
    uiWert : UINT;
    xBekannt : BOOL;
  END_VAR
  VAR_IN_OUT
    aBild : T_VP_ErzeugerBild;
  END_VAR

IF xBekannt THEN
    aBild[uiAdresse] := UINT_TO_WORD(uiWert);
ELSE
    aBild[uiAdresse] := 16#FFFF;
END_IF
VP_SetzeU16 := xBekannt;
END_FUNCTION

FUNCTION VP_SetzeS16 : BOOL
  VAR_INPUT
    uiAdresse : UINT;
    iWert : INT;
    xBekannt : BOOL;
  END_VAR
  VAR_IN_OUT
    aBild : T_VP_ErzeugerBild;
  END_VAR

IF xBekannt THEN
    (* Zweierkomplement: INT_TO_WORD behält das Bitmuster *)
    aBild[uiAdresse] := INT_TO_WORD(iWert);
ELSE
    aBild[uiAdresse] := 16#7FFF;
END_IF
VP_SetzeS16 := xBekannt;
END_FUNCTION

FUNCTION VP_SetzeU32 : BOOL
  VAR_INPUT
    uiAdresse : UINT;
    udiWert : UDINT;
    xBekannt : BOOL;
  END_VAR
  VAR_IN_OUT
    aBild : T_VP_ErzeugerBild;
  END_VAR

IF xBekannt THEN
    aBild[uiAdresse] := UDINT_TO_WORD(SHR(udiWert, 16));
    aBild[uiAdresse + 1] := UDINT_TO_WORD(udiWert AND 16#FFFF);
ELSE
    aBild[uiAdresse] := 16#FFFF;
    aBild[uiAdresse + 1] := 16#FFFF;
END_IF
VP_SetzeU32 := xBekannt;
END_FUNCTION

FUNCTION VP_SetzeS32 : BOOL
  VAR_INPUT
    uiAdresse : UINT;
    diWert : DINT;
    xBekannt : BOOL;
  END_VAR
  VAR_IN_OUT
    aBild : T_VP_ErzeugerBild;
  END_VAR

IF xBekannt THEN
    (* Zweierkomplement über dieselbe Routine wie jeder 32-bit-Wert: DINT_TO_UDINT behält das Bitmuster *)
    VP_SetzeU32(aBild := aBild, uiAdresse := uiAdresse, udiWert := DINT_TO_UDINT(diWert), xBekannt := TRUE);
ELSE
    aBild[uiAdresse] := 16#7FFF;
    aBild[uiAdresse + 1] := 16#FFFF;
END_IF
VP_SetzeS32 := xBekannt;
END_FUNCTION

(* Ein Name: 16 Wörter = 32 Zeichen ISO 8859-1, höherwertiges Byte zuerst, mit 0 aufgefüllt (Vertrag §6). *)
FUNCTION VP_SetzeText : BOOL
  VAR_INPUT
    uiAdresse : UINT;
    sText : STRING(32);
  END_VAR
  VAR_IN_OUT
    aBild : T_VP_ErzeugerBild;
  END_VAR
  VAR
    iLaenge : INT;
    i : INT;
    bHoch : BYTE;
    bNieder : BYTE;
  END_VAR

iLaenge := LEN(sText);
FOR i := 0 TO 15 DO
    bHoch := 0;
    bNieder := 0;
    (* Hinter dem Ende des Texts steht 0, nie ein Rest aus dem Speicher der Zeichenkette *)
    IF 2 * i < iLaenge THEN
        bHoch := sText[2 * i];
    END_IF
    IF 2 * i + 1 < iLaenge THEN
        bNieder := sText[2 * i + 1];
    END_IF
    aBild[uiAdresse + INT_TO_UINT(i)] := SHL(BYTE_TO_WORD(bHoch), 8) OR BYTE_TO_WORD(bNieder);
END_FOR
VP_SetzeText := iLaenge > 0;
END_FUNCTION

(* Ein Bit eines Bitfelds. *)
FUNCTION VP_Bit : WORD
  VAR_INPUT
    xGesetzt : BOOL;
    uiBit : UINT;
  END_VAR

IF xGesetzt THEN
    VP_Bit := SHL(WORD#1, uiBit);
ELSE
    VP_Bit := 0;
END_IF
END_FUNCTION

(* VoltPilot-Bibliothek · Packen, Lesen und Siegel des Koppelbilds Wortfolge wie im Erzeuger-Bild: höherwertiges Wort zuerst; ungültig ist das Typ-Maximum. Auch der Prüfwert 16#01020304 der Quittung geht über VP_KoppelSetzeU32 (Vertrag §1). *)
FUNCTION VP_KoppelSetzeU32 : BOOL
  VAR_INPUT
    uiAdresse : UINT;
    udiWert : UDINT;
  END_VAR
  VAR_IN_OUT
    aQ : T_VP_KoppelQuittung;
  END_VAR

aQ[uiAdresse] := UDINT_TO_WORD(SHR(udiWert, 16));
aQ[uiAdresse + 1] := UDINT_TO_WORD(udiWert AND 16#FFFF);
VP_KoppelSetzeU32 := TRUE;
END_FUNCTION

FUNCTION VP_KoppelSetzeS32 : BOOL
  VAR_INPUT
    uiAdresse : UINT;
    diWert : DINT;
    xBekannt : BOOL;
  END_VAR
  VAR_IN_OUT
    aQ : T_VP_KoppelQuittung;
  END_VAR

IF xBekannt THEN
    (* Zweierkomplement: DINT_TO_UDINT behält das Bitmuster *)
    VP_KoppelSetzeU32(aQ := aQ, uiAdresse := uiAdresse, udiWert := DINT_TO_UDINT(diWert));
ELSE
    aQ[uiAdresse] := 16#7FFF;
    aQ[uiAdresse + 1] := 16#FFFF;
END_IF
VP_KoppelSetzeS32 := xBekannt;
END_FUNCTION

(* Ein 32-bit-Wert aus zwei Wörtern des Wunschs, höherwertiges Wort zuerst. *)
FUNCTION VP_KoppelLiesU32 : UDINT
  VAR_INPUT
    uiAdresse : UINT;
  END_VAR
  VAR_IN_OUT
    aW : T_VP_KoppelWunsch;
  END_VAR

VP_KoppelLiesU32 := SHL(WORD_TO_UDINT(aW[uiAdresse]), 16) OR WORD_TO_UDINT(aW[uiAdresse + 1]);
END_FUNCTION

(* Ein Wort in die CRC-16/MODBUS (Polynom 16#A001 gespiegelt): erst das höherwertige Byte. *)
FUNCTION VP_KoppelCrcWort : WORD
  VAR_INPUT
    wCrc : WORD;
    wWort : WORD;
  END_VAR
  VAR
    wC : WORD;
    wByte : WORD;
    k : INT;
    i : INT;
  END_VAR

wC := wCrc;
FOR k := 0 TO 1 DO
    IF k = 0 THEN
        wByte := SHR(wWort, 8);
    ELSE
        wByte := wWort AND 16#00FF;
    END_IF
    wC := wC XOR wByte;
    FOR i := 1 TO 8 DO
        IF (wC AND 16#0001) <> 0 THEN
            wC := SHR(wC, 1) XOR 16#A001;
        ELSE
            wC := SHR(wC, 1);
        END_IF
    END_FOR
END_FOR
VP_KoppelCrcWort := wC;
END_FUNCTION

(* Siegel des Wunschs: über die Wörter 0..14 und 16..63 (Vertrag §8). *)
FUNCTION VP_KoppelSiegelW : WORD
  VAR_IN_OUT
    aW : T_VP_KoppelWunsch;
  END_VAR
  VAR
    wC : WORD;
    i : UINT;
  END_VAR

wC := 16#FFFF;
FOR i := 0 TO 63 DO
    IF i <> 15 THEN
        wC := VP_KoppelCrcWort(wCrc := wC, wWort := aW[i]);
    END_IF
END_FOR
VP_KoppelSiegelW := wC;
END_FUNCTION

(* Siegel der Quittung: über die Wörter 1000..1018 und 1020..1115, hier 0..18 und 20..115. *)
FUNCTION VP_KoppelSiegelQ : WORD
  VAR_IN_OUT
    aQ : T_VP_KoppelQuittung;
  END_VAR
  VAR
    wC : WORD;
    i : UINT;
  END_VAR

wC := 16#FFFF;
FOR i := 0 TO 115 DO
    IF i <> 19 THEN
        wC := VP_KoppelCrcWort(wCrc := wC, wWort := aQ[i]);
    END_IF
END_FOR
VP_KoppelSiegelQ := wC;
END_FUNCTION

(* VoltPilot-Bibliothek · Packfunktion des WAGO-Bilds Jeder 32-bit-Wert geht über VP_WagoSetze32 ins Bild - auch der Prüfwert 16#01020304 (Vertrag §3): er bestätigt der Box die Wortfolge nur, wenn er durch dieselbe Routine geht wie die Messwerte. Wortfolge (Parameter je Anlage, Vertrag §2): FALSE = höherwertiges Wort zuerst ("big"), TRUE = niederwertiges zuerst ("little"). Innerhalb eines Worts gilt die Modbus-Byte-Reihenfolge. *)
FUNCTION VP_WagoSetze32 : BOOL
  VAR_INPUT
    uiAdresse : UINT;
    dwWert : DWORD;
    xLittle : BOOL;
  END_VAR
  VAR_IN_OUT
    aBild : T_VP_WagoBild;
  END_VAR

IF xLittle THEN
    aBild[uiAdresse] := DWORD_TO_WORD(dwWert AND 16#FFFF);
    aBild[uiAdresse + 1] := DWORD_TO_WORD(SHR(dwWert, 16));
ELSE
    aBild[uiAdresse] := DWORD_TO_WORD(SHR(dwWert, 16));
    aBild[uiAdresse + 1] := DWORD_TO_WORD(dwWert AND 16#FFFF);
END_IF
VP_WagoSetze32 := TRUE;
END_FUNCTION

(* VoltPilot-Vorlage PV (Entscheid E3 = A): Anlagenprogramm einer PV-Anlage mit bis zu 10 Wechselrichtern, das den Wunsch der Box annimmt. Der Fachbetrieb passt die mit ANPASSEN markierten Zeilen an: Eingänge der Anlage, Vorgabe des Netzbetreibers, Ausgabe an die Wechselrichter. Stellplatz 1: limit_w auf die ganze Erzeugung, Band 0 W bis Nennleistung. Vorrang bleibt im Anlagenprogramm: wirksam ist das Kleinste aus Nennleistung, Grenze des Netzbetreibers und gültigem Wunsch. Bestimmt der Netzbetreiber statt des Wunschs, meldet die Rückmeldung "überstimmt" und das Angebot grund_vorrang. Ohne gültigen Wunsch (Box aus, Frist vorbei, Schlüsselschalter auf Ort) fährt die Anlage mit ihren eigenen Werten. Die wirksame Grenze steht im Erzeuger-Bild (p_grenze_w); bestimmt der Wunsch sie, nennt quelle_p keine Stelle (0) - wer stellt, sagt die Quittung des Koppelbilds (Erzeuger-Bild bleibt 1.0). *)
PROGRAM PLC_PRG
  VAR
    udiSteuerungId : UDINT := 1;
    uiProgrammstand : UINT := 2611;
    uiTeAnzahl : UINT := 3;
    auiNennKw : ARRAY[1..10] OF UINT;
    xSchluesselFern : BOOL := TRUE;
    xHandOrt : BOOL;
    xStoerung : BOOL;
    xNbVorgabe : BOOL;
    uiNbZehntelProzent : UINT := 1000;
    audiSollW : ARRAY[1..10] OF UDINT;
    fbBild : FB_VP_ErzeugerBild;
    fbKoppel : FB_VP_Koppelbild;
    stAnlage : ST_VP_ErzeugerAnlage;
    stNb : ST_VP_ErzeugerNetzbetreiber;
    stDv : ST_VP_ErzeugerDirektvermarkter;
    stWirkung : ST_VP_ErzeugerWirkung;
    astEinheit : ARRAY[1..10] OF ST_VP_ErzeugerEinheit;
    aAngebot : ARRAY[1..8] OF ST_VP_Angebot;
    aRueck : ARRAY[1..8] OF ST_VP_Rueckmeldung;
    udiNennW : UDINT;
    diNenn : DINT;
    diNb : DINT;
    diGrenze : DINT;
    n : UINT;
  END_VAR

(* --- Nennleistung -------------------------------------------------------------------------- *)
udiNennW := 0;
FOR n := 1 TO uiTeAnzahl DO
    udiNennW := udiNennW + UINT_TO_UDINT(auiNennKw[n]) * 1000;
END_FOR
diNenn := UDINT_TO_DINT(udiNennW);

(* --- Angebot: Stellplatz 1 begrenzt die ganze Erzeugung ------------------------------------ *)
aAngebot[1].uiArt := 1;    (* limit_w *)
aAngebot[1].uiZiel := 1;   (* erzeugung_gesamt *)
aAngebot[1].diMin := 0;
aAngebot[1].diMax := diNenn;
aAngebot[1].xBereit := NOT xStoerung;
aAngebot[1].xGrundStoerung := xStoerung;

fbKoppel(udiSteuerungId := udiSteuerungId, xFernsteuerungFrei := xSchluesselFern, xHandOrt := xHandOrt,
    aAngebot := aAngebot, aRueckmeldung := aRueck, aWunschRegister := GVL_VoltPilot.aKoppelWunsch,
    aQuittungRegister := GVL_VoltPilot.aKoppelQuittung);

(* --- Vorrang: zuerst der Netzbetreiber, dann der Wunsch ------------------------------------ *)
diNb := diNenn;
IF xNbVorgabe THEN
    diNb := MIN(diNenn, UDINT_TO_DINT(udiNennW * UINT_TO_UDINT(uiNbZehntelProzent) / 1000));
END_IF
diGrenze := diNb;
IF fbKoppel.aWunsch[1].xGilt THEN
    diGrenze := MIN(diGrenze, fbKoppel.aWunsch[1].diWert);
END_IF
aRueck[1].diWirksam := diGrenze;
aRueck[1].xWirksamBekannt := diGrenze < diNenn;
aRueck[1].xUeberstimmt := fbKoppel.aWunsch[1].xGilt AND diNb < fbKoppel.aWunsch[1].diWert;
aAngebot[1].xGrundVorrang := diNb < diNenn;

(* --- Ausgabe: die Grenze nach Nennleistung auf die Wechselrichter ------------------------- *)
FOR n := 1 TO uiTeAnzahl DO
    IF udiNennW > 0 THEN
        audiSollW[n] := DINT_TO_UDINT(diGrenze) / 1000 * UINT_TO_UDINT(auiNennKw[n]) * 1000 / (udiNennW / 1000);
    END_IF
    astEinheit[n].xSollwertGueltig := TRUE;
    astEinheit[n].udiPSollW := audiSollW[n];
    astEinheit[n].uiArt := 1;
    astEinheit[n].uiNennKw := auiNennKw[n];
END_FOR

(* --- Erzeuger-Bild: was gilt und wer es bestimmt ------------------------------------------- *)
stAnlage.uiInstalliertKw := UDINT_TO_UINT(udiNennW / 1000);
stAnlage.xHandOrt := xHandOrt;
stAnlage.xSammelstoerung := xStoerung;
stNb.uiKanal := 3;
stNb.xVorgabeGueltig := xNbVorgabe;
stNb.uiPZehntelProzent := uiNbZehntelProzent;
stWirkung.xGueltig := TRUE;
stWirkung.udiGrenzeW := DINT_TO_UDINT(diGrenze);
IF diNb < diNenn AND diNb <= diGrenze THEN
    stWirkung.uiQuelle := 1;   (* netzbetreiber *)
ELSE
    stWirkung.uiQuelle := 0;   (* keine Stelle des Erzeuger-Bilds; der Wunsch steht in der Quittung *)
END_IF
fbBild(udiSteuerungId := udiSteuerungId, uiProgrammstand := uiProgrammstand, uiAnlagenart := 1,
    uiTeAnzahl := uiTeAnzahl, stAnlage := stAnlage, stNetzbetreiber := stNb, stDirektvermarkter := stDv,
    stWirkung := stWirkung, astEinheit := astEinheit, xMitNamen := FALSE, aBild := GVL_VoltPilot.aErzeugerBild);
END_PROGRAM
